Fanuc KAREL source: KC00012.KL

PROGRAM KC00012
%NOLOCKGROUP
%ENVIRONMENT PBQMGR
VAR
  I: INTEGER
  J: INTEGER
  K: INTEGER
  R: REAL
  B: BOOLEAN
  S: STRING[80]
  T: STRING[80]
  P: PATH
  Q: PATH
  QT: QUEUE_TYPE
  AI: ARRAY[8] OF INTEGER
  AB: ARRAY[244] OF BYTE
BEGIN
  COPY_QUEUE(QT,AI,I,J,AI,K,I)
END KC00012
